(* IEC 61131-3 sources: Versio-VersionControlSystem/fixtures/projects/RefrigeratorControl/Device/Plc Logic/Application/Library/Alarm/GVLs, 1 file *)

(* ---- GVL_Alarm.gvl.st ---- *)
{attribute 'qualified_only'}
VAR_GLOBAL
	AlarmConstant : DINT := 3;
END_VAR
